(* IEC 61131-3 sources: JingjiangArm/moonboxpro_arm_8.4/Application/Application/任务列表/TensionTask/电机运动/MotionCtl_Trap, 5 files *)

(* ---- StMotorParam_Trap.st ---- *)
(*@CES
Name=StMotorParam_Trap
Type=Gvl
TypeGuid=2db5746d-d284-4425-9f7f-2663a34b0ebc
Guid=895de25e-1961-43a4-b404-7adc5138347b
HasDeclaration=True
HasImplementation=False
*)
{DECLARATION}
TYPE StMotorParam_Trap ://点位轴和龙门轴的参数
STRUCT
	iAxisId: INT;
	iCoreId: INT;
	iStationId: INT;
	iUnitId : INT;
	iMoveStep: INT;
	xMoveRev: BOOL;
	xMoveEn: BOOL;
	uiAxisNum: UINT;(*减速比分子*)
	uiAxisDen: UINT;(*减速比分母*)
	liTargetPos: LINT;(*点位目标位置*)
	udiTargetVel: UDINT;
	rScrewPitch_: REAL;(*螺距*)
END_STRUCT
END_TYPE

{IMPLEMENTATION}

(* ---- KS_FB_AxisPosCtl_Trap.st ---- *)
(*@CES
Name=KS_FB_AxisPosCtl_Trap
Type=FunctionBlock
TypeGuid=6f9dac99-8de1-4efc-8465-68ac443b7d08
Guid=53966cce-5ce5-480b-a4cc-b0ff05bfaf84
HasDeclaration=True
HasImplementation=True
*)
{DECLARATION}
FUNCTION_BLOCK KS_FB_AxisPosCtl_Trap
VAR_INPUT
	i_xEn: BOOL;
	i_iGrpId: INT;
	i_iGrpUnitNum_Pu : INT;
	i_aiGrpUnitList: ARRAY [1..MAX_UNIT_NUM] OF INT;
	i_iGrpTrapMotion_Num: INT;
	i_aiGrpTrapMotion_StdList: ARRAY [1..MAX_STATION_NUM] OF INT;
	i_pstStSysParam: POINTER TO StSysParam;
	i_pastStMotorParam_Trap: POINTER TO ARRAY [1..MAX_STATION_NUM] OF StMotorParam_Trap;

	i_xHorManuCtrl:BOOL;(*界面横向手动修正功能*)

	//2026.01.28.173520 | + | 横向伺服控制
	i_alrTarp_EncPos						: ARRAY [1..MAX_UNIT_NUM] OF LREAL;//横向点位轴的编码器位置
	i_pastStIOMap_AxisBasic					: POINTER TO ARRAY [1..MAX_UNIT_NUM] OF StIOMap_Axis_FE; (*基础io|*)
	i_pastStAxisRapidAdjProf_H				: POINTER TO ARRAY [1..MAX_UNIT_NUM] OF StAxisRapidAdjProf_H;(*纵向快速对版|*)

	i_paxLimit_Left_Wr 						: POINTER TO ARRAY [1..MAX_UNIT_NUM] OF BOOL;
 	i_paxLimit_Right_Wr 					: POINTER TO ARRAY [1..MAX_UNIT_NUM] OF BOOL;
	i_paxLimit_Left_WrClr 					: POINTER TO ARRAY [1..MAX_UNIT_NUM] OF BOOL;
 	i_paxLimit_Right_WrClr 					: POINTER TO ARRAY [1..MAX_UNIT_NUM] OF BOOL;

	//新增拿横向编码器 2026.05.09.104451
	i_pastStGetMotionSts			: POINTER TO ARRAY [1..MAX_STATION_NUM] OF StGetMotionSts;
	i_pstStSysStationInf			:POINTER TO StSysStationInf;
	i_pstStSysGantryAxisInf 		:POINTER TO StSysGantryAxisInf;
	i_pastStAxisIdListInf 			:POINTER TO ARRAY [1..128] OF StAxisIdListInf;
END_VAR
VAR_OUTPUT
END_VAR
VAR
	iN: INT;
	iAxisId: INT;
	iTypeId: INT;
	iUnitId: INT;
	iCoreId: INT;
	pstStGrpParam_Save: POINTER TO StGrpParam_Save;
	pstStGrpParam_UnSave: POINTER TO StGrpParam_UnSave;

	//2026.01.28.173520 | + | 横向伺服控制
	fbKS_FB_HorzCtl_Driver : KS_FB_HorzCtl_Driver;

	alrTotalAdjust_Horz : ARRAY [1..MAX_UNIT_NUM] OF LREAL;
END_VAR

{IMPLEMENTATION}
IF i_xEn THEN
	IF (i_iGrpId=1 OR i_iGrpId=2) AND
		i_iGrpUnitNum_Pu>=1 AND i_iGrpUnitNum_Pu<=MAX_UNIT_NUM AND
		i_iGrpTrapMotion_Num>=1 AND i_iGrpTrapMotion_Num<= MAX_STATION_NUM AND
		i_pstStSysParam<>0 AND
		i_pastStMotorParam_Trap<>0 THEN
		pstStGrpParam_Save:= ADR(i_pstStSysParam^.astStGrpParam_Save[i_iGrpId]);
		pstStGrpParam_UnSave:= ADR(i_pstStSysParam^.astStGrpParam_UnSave[i_iGrpId]);

		//2026.01.28.173520 | + | 横向伺服控制
		fbKS_FB_HorzCtl_Driver(
			i_xEn:= TRUE,//(pstStGrpParam_UnSave^.xFlag_Print OR i_pstStSysParam^.astStGrpParam_Save[i_iGrpId].xEnaTestARC_Ink (*空转测试使能*)) AND g_stStSysParam.stStSysParam_Save.byHorzCtlMode=3,
			i_iGrpId:= i_iGrpId,
			i_iGrpAxisNum_Pu:= i_iGrpUnitNum_Pu,
			i_pstStSysParam:= i_pstStSysParam,
			i_pastStIOMap_AxisBasic:= i_pastStIOMap_AxisBasic,
			i_lrVel_HorzAdjust:= REAL_TO_LREAL(i_pstStSysParam^.astStGrpParam_Save[i_iGrpId].rVel_HorzdAdj),
			i_lrVel_HorzPreRegister:=  REAL_TO_LREAL(i_pstStSysParam^.astStGrpParam_Save[i_iGrpId].rVel_HorzPreRegister),
			i_xFlag_Estop:= pstStGrpParam_UnSave^.xFlag_EStop,
			i_xFlag_Stop:= pstStGrpParam_UnSave^.xFlag_Stop,
			i_iCycleTime_Plc:= gc_TENSION_TSK_CYCLE_TIME,
			i_pastStAxisRapidAdjProf_H:= i_pastStAxisRapidAdjProf_H,
			i_alrTarp_EncPos:= i_alrTarp_EncPos,
			i_paxLimit_Left_Wr:= i_paxLimit_Left_Wr,
			i_paxLimit_Right_Wr:= i_paxLimit_Right_Wr,
			i_paxLimit_Left_WrClr:= i_paxLimit_Left_WrClr,
			i_paxLimit_Right_WrClr:= i_paxLimit_Right_WrClr,
			i_xHorManuCtrl:= i_xHorManuCtrl,
			i_aiGrpTrapMotion_StdList:=i_aiGrpTrapMotion_StdList,
			i_pastStGetMotionSts:=i_pastStGetMotionSts,
			i_pstStSysStationInf:=i_pstStSysStationInf,
			i_pstStSysGantryAxisInf :=i_pstStSysGantryAxisInf,
			i_pastStAxisIdListInf :=i_pastStAxisIdListInf,
			o_xEno=> ,
			o_iErNo=> ,
			o_alrTotalAdjust_Horz=> alrTotalAdjust_Horz);

		FOR iN:=1 TO i_iGrpTrapMotion_Num BY 1 DO
			i_pastStMotorParam_Trap^[iN].liTargetPos := LREAL_TO_LINT(alrTotalAdjust_Horz[iN]*
						i_pstStSysParam^.astStUnitParam_Save[iN].uiNum_Horz*
						GC_LRMOTORPPR_TRAP/
						i_pstStSysParam^.astStUnitParam_Save[iN].rScrewPitch_Horz/
						i_pstStSysParam^.astStUnitParam_Save[iN].uiDen_Horz/1000.0);
			i_pastStMotorParam_Trap^[iN].udiTargetVel := LREAL_TO_UDINT(i_pstStSysParam^.astStGrpParam_Save[i_iGrpId].rVel_HorzdAdj*
						i_pstStSysParam^.astStUnitParam_Save[iN].uiNum_Horz*
						GC_LRMOTORPPR_TRAP/
						i_pstStSysParam^.astStUnitParam_Save[iN].rScrewPitch_Horz/
						i_pstStSysParam^.astStUnitParam_Save[iN].uiDen_Horz/1000.0);
		END_FOR
	END_IF
ELSE
	;
END_IF

(* ---- KS_FB_HorzCtl_Driver.st ---- *)
(*@CES
Name=KS_FB_HorzCtl_Driver
Type=FunctionBlock
TypeGuid=6f9dac99-8de1-4efc-8465-68ac443b7d08
Guid=da6152f2-d53e-407a-9477-cd718a7d485f
HasDeclaration=True
HasImplementation=True
*)
{DECLARATION}
FUNCTION_BLOCK KS_FB_HorzCtl_Driver
VAR_INPUT
	i_xEn: BOOL;(*使能*)
	i_iGrpId: INT;
	i_iGrpAxisNum_Pu: INT; (*色组轴数*)
	i_pstStSysParam:POINTER TO StSysParam;(*系参数*)
	i_pastStIOMap_AxisBasic					: POINTER TO ARRAY [1..MAX_UNIT_NUM] OF StIOMap_Axis_FE; (*基础io|*)
	i_lrVel_HorzAdjust		: LREAL;(*mm/s; um/ms; 横向调整速度|*)
	i_lrVel_HorzPreRegister		: LREAL;(*mm/s;横向预套准速度|*)
	(*2023.3.8.114628*)
	i_xFlag_Estop							: BOOL;(*急停标志*)
	i_xFlag_Stop							: BOOL;(*停机标志*)
	i_iCycleTime_Plc						: INT;
	i_pastStAxisRapidAdjProf_H				: POINTER TO ARRAY [1..MAX_UNIT_NUM] OF StAxisRapidAdjProf_H;(*纵向快速对版|*)
	i_alrTarp_EncPos						: ARRAY [1..MAX_UNIT_NUM] OF LREAL;//横向点位轴的编码器位置
	i_paxLimit_Left_Wr 						: POINTER TO ARRAY [1..MAX_UNIT_NUM] OF BOOL;
 	i_paxLimit_Right_Wr 					: POINTER TO ARRAY [1..MAX_UNIT_NUM] OF BOOL;
	i_paxLimit_Left_WrClr 						: POINTER TO ARRAY [1..MAX_UNIT_NUM] OF BOOL;
 	i_paxLimit_Right_WrClr 					: POINTER TO ARRAY [1..MAX_UNIT_NUM] OF BOOL;
	i_xHorManuCtrl:BOOL;(*界面横向手动修正功能*)
//	i_arStep_Horz			:POINTER TO ARRAY [1..MAX_UNIT_NUM] OF REAL;
//2026.05.09.100428 新增横向标定功能
	i_aiGrpTrapMotion_StdList: ARRAY [1..MAX_STATION_NUM] OF INT;
	i_pastStGetMotionSts: POINTER TO ARRAY [1..MAX_STATION_NUM] OF StGetMotionSts;
	i_pstStSysStationInf			:POINTER TO StSysStationInf;
	i_pstStSysGantryAxisInf 		:POINTER TO StSysGantryAxisInf;
	i_pastStAxisIdListInf :POINTER TO ARRAY [1..128] OF StAxisIdListInf;
END_VAR
VAR_OUTPUT
	o_xEno: BOOL;
	o_iErNo: INT;(*0成功\-1参数失败|*)
	o_alrTotalAdjust_Horz: ARRAY [1..MAX_UNIT_NUM] OF LREAL;(*横向调整量*)

END_VAR
VAR
	iN: INT;
	xInit: BOOL;
	iAxisId: INT;
	pstStGrpParam_Save: POINTER TO StGrpParam_Save;
	pstStGrpParam_UnSave: POINTER TO StGrpParam_UnSave;

	pstStUnitParam_Save: POINTER TO StUnitParam_Save;
	pstStUnitParam_UnSave: POINTER TO StUnitParam_UnSave;
	pstStRSV_UnitParam_Save: POINTER TO StRSV_UnitParam_Save;
	pstStRSV_UnitParam_UnSave: POINTER TO StRSV_UnitParam_UnSave;
	(*横向运动相关变量都使用操作侧和传动侧变量重新赋值@2023.3.8.104853*)
	axHorMovingBtn_M: ARRAY [1..MAX_UNIT_NUM] OF BOOL;(*横向操作侧运动按钮*)
	axHorMovingBtn_G: ARRAY [1..MAX_UNIT_NUM] OF BOOL;(*横向传动侧运动按钮*)
	axHorMovingLimit_M: ARRAY [1..MAX_UNIT_NUM] OF BOOL;(*横向操作侧运动限位*)
	axHorMovingLimit_G: ARRAY [1..MAX_UNIT_NUM] OF BOOL;(*横向传动侧运动限位*)
	axHorMoving_M: ARRAY [1..MAX_UNIT_NUM] OF BOOL;(*横向操作侧运动*)
	axHorMoving_G: ARRAY [1..MAX_UNIT_NUM] OF BOOL;(*横向传动侧运动*)

	lrAdjustVel_:LREAL;(*每个周期调整的量|这里还是mm/s，需要转化为*)
	alrTotalAdjust_Horz: ARRAY [1..MAX_UNIT_NUM] OF LREAL;(*横向调整量*)
	adwTotalTimes_CW_AxisHorzManu: ARRAY [1..MAX_UNIT_NUM] OF DWORD := [MAX_UNIT_NUM(0)];
	adwTotalTimes_CCW_AxisHorzManu: ARRAY [1..MAX_UNIT_NUM] OF DWORD := [MAX_UNIT_NUM(0)];

	wHorzMotorDir: WORD;(*.0 |正转方向
					.1|反转方向*)
	awPreHorzMotorDir: ARRAY [1..MAX_UNIT_NUM] OF WORD;
	axHorzMotorStart_Delay: ARRAY [1..MAX_UNIT_NUM] OF BOOL;(*横向启动延时标志*)
	axHorzMotorStart_DelayDne: ARRAY [1..MAX_UNIT_NUM] OF BOOL;(*横向启动延时完成*)
	auiHorzMotorStart_Count: ARRAY [1..MAX_UNIT_NUM] OF UINT;(*启动延时计时变量*)
	iHorzMotorStart_DelayTime_MS: INT:=0;(*启动的延时时间ms*)

	axStopManuMove_Horz: ARRAY  [1..MAX_UNIT_NUM] OF BOOL;
	lrLimit_Left:LREAL;
	lrLimit_Right:LREAL;
	xLimit_LeftTemp:BOOL;
	xLimit_RightTemp:BOOL;
	xLimit_Left:BOOL;
	xLimit_Right:BOOL;
	lrAbsPosHorz:LREAL;
	iRtn:INT;
	xAxisRev:BOOL;

	//2026.05.09.170157 | + | 增加正反流向
	xMachineIsRev : BOOL;
END_VAR

{IMPLEMENTATION}
o_xEno:= i_xEn;
o_iErNo:= 0;
IF i_xEn THEN
	IF (i_iGrpAxisNum_Pu>=1 AND i_iGrpAxisNum_Pu<=MAX_UNIT_NUM) AND(*系的色组数量有效|*)
		i_pstStSysParam<>0 AND(*参数有效|*)
		i_pastStIOMap_AxisBasic<>0 AND
		i_paxLimit_Left_Wr<>0 AND
		i_paxLimit_Right_Wr<>0 THEN

		pstStGrpParam_Save :=  ADR(i_pstStSysParam^.astStGrpParam_Save[i_iGrpId]);
		pstStGrpParam_UnSave :=  ADR(i_pstStSysParam^.astStGrpParam_UnSave[i_iGrpId]);
		//初始化输出调整量为当前规划位置
// 		IF NOT xInit THEN
// 			xInit:= TRUE;
// 			FOR iN:=1 TO i_iGrpAxisNum_Pu BY 1 DO
// 				alrTotalAdjust_Horz[iN]:= i_alrTarp_PrfPos[iN];
// 			END_FOR
// 		END_IF

		//2026.05.09.170157 | + | 增加正反流向
		xMachineIsRev := TRUE;

		IF NOT xInit THEN
			xInit:= TRUE;
			FOR iN:=1 TO i_iGrpAxisNum_Pu BY 1 DO
				alrTotalAdjust_Horz[iN]:= 0;
			END_FOR
		END_IF
		(*2023.3.8.114227 将函数KS_FB_AxisHorAdj中的代码移植到此处*)
		FOR iN:= 1 TO i_iGrpAxisNum_Pu BY 1 DO
			iAxisId:= iN;
			pstStUnitParam_Save:= ADR(i_pstStSysParam^.astStUnitParam_Save[iAxisId]);
			pstStUnitParam_UnSave:= ADR(i_pstStSysParam^.astStUnitParam_UnSave[iAxisId]);

			pstStRSV_UnitParam_Save := ADR(i_pstStSysParam^.astStRSV_UnitParam_Save[iAxisId]);
			pstStRSV_UnitParam_UnSave := ADR(i_pstStSysParam^.astStRSV_UnitParam_UnSave[iAxisId]);

			(*处理一下限位*)
			(*限位赋值*)
			IF pstStGrpParam_UnSave^.xIsDebugMode_Machine AND pstStGrpParam_UnSave^.xFlag_Stop THEN//调试模式
				//记录一下横向限位
				IF i_paxLimit_Left_Wr^[iAxisId] THEN
					i_paxLimit_Left_Wr^[iAxisId]:= FALSE;
					//2026.05.09.100428 新增横向标定功能 Hou.N
					iRtn := GTN_RN_ReadAbsEncPos(cardIndex:= 1, stationPhyId:=i_aiGrpTrapMotion_StdList[iAxisId], encoder:= 1, pPos:= ADR(lrAbsPosHorz));
					g_liAbsPosTrap := LREAL_TO_LINT(lrAbsPosHorz);
					xAxisRev := pstStUnitParam_UnSave^.xMotRev_Horiz_;
					iRtn := KS_SetTrapCoordinate(
							i_xEn:= TRUE,
							i_iTarget_Num:= 1,
							i_paiTargetStationList:= ADR(i_aiGrpTrapMotion_StdList[iAxisId]),
							i_paliABSEncPos:= ADR(g_liAbsPosTrap),
							i_paxAxisRev:= ADR(xAxisRev),
							i_pastStAxisIdListInf:= i_pastStAxisIdListInf,
							i_pastStGetMotionSts:= i_pastStGetMotionSts,
							i_pstStSysStationInf := i_pstStSysStationInf,
							i_pstStSysGantryAxisInf := i_pstStSysGantryAxisInf,
							ADR(g_alrCurrentAbsPos_Trap));
					i_pstStSysParam^.astStRSV_UnitParam_Save[iAxisId].liABSPos_Trap:= g_liAbsPosTrap;
					pstStRSV_UnitParam_Save^.lrLimit_Left:= 1;
				END_IF

				IF i_paxLimit_Right_Wr^[iAxisId] THEN
					i_paxLimit_Right_Wr^[iAxisId]:= FALSE;
					pstStRSV_UnitParam_Save^.lrLimit_Right:= i_alrTarp_EncPos[iAxisId];
				END_IF
				IF 	i_paxLimit_Left_WrClr^[iAxisId] THEN
					i_paxLimit_Left_WrClr^[iAxisId] := FALSE;
					pstStRSV_UnitParam_Save^.lrLimit_Left := 0;
					i_pstStSysParam^.astStRSV_UnitParam_Save[iAxisId].liABSPos_Trap:=0;
				END_IF
				IF 	i_paxLimit_Right_WrClr^[iAxisId] THEN
					i_paxLimit_Right_WrClr^[iAxisId] := FALSE;
					pstStRSV_UnitParam_Save^.lrLimit_Right := 0;
				END_IF
			ELSE
				i_paxLimit_Left_Wr^[iAxisId]:= FALSE;
				i_paxLimit_Right_Wr^[iAxisId]:= FALSE;
				i_paxLimit_Left_WrClr^[iAxisId]:= FALSE;
				i_paxLimit_Right_WrClr^[iAxisId]:= FALSE;
			END_IF
			lrLimit_Left:= pstStRSV_UnitParam_Save^.lrLimit_Left;
			lrLimit_Right:= pstStRSV_UnitParam_Save^.lrLimit_Right;
			xLimit_LeftTemp:=i_pastStIOMap_AxisBasic^[iAxisId].i_xPosLimit_Left;
			xLimit_RightTemp:=i_pastStIOMap_AxisBasic^[iAxisId].i_xPosLimit_Right;

			IF lrLimit_Left=0 THEN(*未有软限位|按照最远距离*);

			ELSE(*存在软限位|限位标志取接近开关和位置值的or*)
				IF pstStUnitParam_UnSave^.xMotRev_Horiz_ THEN
					xLimit_LeftTemp:=xLimit_LeftTemp OR
									(lrLimit_Left<i_alrTarp_EncPos[iAxisId]);
				ELSE
					xLimit_LeftTemp:=xLimit_LeftTemp OR
									(lrLimit_Left<i_alrTarp_EncPos[iAxisId]);
				END_IF
			END_IF
			IF lrLimit_Right=0 THEN(*未有软限位|按照最远距离*);
			ELSE(*存在软限位|限位标志取接近开关和位置值的or*)
				IF pstStUnitParam_UnSave^.xMotRev_Horiz_ THEN
					xLimit_RightTemp:=xLimit_RightTemp OR
								(lrLimit_Right>i_alrTarp_EncPos[iAxisId]);
				ELSE
					xLimit_RightTemp:=xLimit_RightTemp OR
								(lrLimit_Right>i_alrTarp_EncPos[iAxisId]);

				END_IF
			END_IF

			(*手动左右取反*)(*bai.zy|2023.12.18.161830|feida取反*)
			xLimit_Left:=xLimit_RightTemp;
			xLimit_Right:=xLimit_LeftTemp;
			(*
			IF xMachineIsRev THEN
				xLimit_Left:=xLimit_RightTemp;
				xLimit_Right:=xLimit_LeftTemp;
				IF pstStUnitParam_UnSave^.xMotRev_Horiz_ THEN
					xLimit_Left:=xLimit_LeftTemp;
					xLimit_Right:=xLimit_RightTemp;
				END_IF
			ELSE
				xLimit_Left:=xLimit_LeftTemp;
				xLimit_Right:=xLimit_RightTemp;
				IF pstStUnitParam_UnSave^.xMotRev_Horiz_ THEN
					xLimit_Left:=xLimit_LeftTemp;
					xLimit_Right:=xLimit_RightTemp;
				END_IF
			END_IF
			*)
//2026.01.28.152311 | + | 界面上的限位提示，先不要了
// 			g_axLimit_Left_Wr_HMI[iN]:= xLimit_Left;
// 			g_axLimit_Right_Wr_HMI[iN]:= xLimit_Right;
			(*处理横向开关相关@2023.3.8.104924*)
			(*和运动方向关联@伺服正转(正手机)-左对应操作侧#先不关心反印时候的方向变化问题
						    @伺服反转(反手机)-左对应传动侧#先不关心反印时候的方向变化问题*)

//			IF pstStUnitParam^.xMotRev_PrnRoller THEN(*正转*)
				axHorMovingBtn_M[iAxisId]:=i_pastStIOMap_AxisBasic^[iAxisId].i_xMove_Left;
				axHorMovingBtn_G[iAxisId]:=i_pastStIOMap_AxisBasic^[iAxisId].i_xMove_Right;

				axHorMovingLimit_M[iAxisId]:=xLimit_Left;
				axHorMovingLimit_G[iAxisId]:=xLimit_Right;
(*			ELSE(*反转*)
				axHorMovingBtn_M[iAxisId]:=pstStIOMap_Axis_FLEXO^.i_xMove_Right;
				axHorMovingBtn_G[iAxisId]:=pstStIOMap_Axis_FLEXO^.i_xMove_Left;

				IF i_pstStSysParam^.dwControlComplexBits.17 THEN
					(*使用左右限位*)
					axHorMovingLimit_M[iAxisId]:=xLimit_Right;
					axHorMovingLimit_G[iAxisId]:=xLimit_Left;
				ELSE
					(*使用正转(操作侧)反转(传动侧)限位*)
					axHorMovingLimit_M[iAxisId]:=xLimit_Left;
					axHorMovingLimit_G[iAxisId]:=xLimit_Right;
				END_IF
			END_IF
*)

			IF i_pastStIOMap_AxisBasic^[iAxisId].o_xRel_Press OR (NOT i_pastStIOMap_AxisBasic^[iAxisId].i_xHorzMotor_FastSpd) THEN
			(*快调/慢调处理*)
				lrAdjustVel_:= i_lrVel_HorzAdjust;
			ELSE
				lrAdjustVel_:= i_lrVel_HorzPreRegister;
			END_IF

			(*2019.5.15.170941|niu.j|急停清零横向调整量*)
			IF pstStGrpParam_UnSave^.xFlag_EStoping OR pstStGrpParam_UnSave^.xFlag_Estop THEN
				pstStUnitParam_UnSave^.alrTotalAdjustVal_Auto_vh[2]:= 0;
				pstStUnitParam_UnSave^.alrTotalAdjustVal_ManuFine_vh[2]:= 0;
				pstStUnitParam_UnSave^.alrTotalAdjustVal_Rapid_vh[2]:= 0;
			END_IF

			IF (pstStUnitParam_Save^.dwFlag_Ctl.0 AND pstStUnitParam_Save^.dwFlag_Sts.1) THEN
				IF ABS(pstStUnitParam_UnSave^.alrTotalAdjustVal_Auto_vh[2])>0 THEN
					IF pstStUnitParam_UnSave^.alrTotalAdjustVal_Auto_vh[2]>0 THEN
						(*正向*)
						alrTotalAdjust_Horz[iAxisId]:= alrTotalAdjust_Horz[iAxisId]+pstStUnitParam_UnSave^.alrTotalAdjustVal_Auto_vh[2];
						pstStUnitParam_UnSave^.alrTotalAdjustVal_Auto_vh[2]:= 0;
						pstStUnitParam_UnSave^.axCurCycleAdjustVal_Auto_done_vh[2]:= FALSE;
						axHorMoving_M[iAxisId]:= TRUE;(*操作侧*)
						axHorMoving_G[iAxisId]:= FALSE;(*传动侧*)
					ELSE
						(*反向*)
						alrTotalAdjust_Horz[iAxisId]:= alrTotalAdjust_Horz[iAxisId]+pstStUnitParam_UnSave^.alrTotalAdjustVal_Auto_vh[2];
						pstStUnitParam_UnSave^.alrTotalAdjustVal_Auto_vh[2]:= 0;
						pstStUnitParam_UnSave^.axCurCycleAdjustVal_Auto_done_vh[2]:= FALSE;
						axHorMoving_G[iAxisId]:= TRUE;(*传动侧*)
						axHorMoving_M[iAxisId]:= FALSE;(*操作侧*)
					END_IF
				ELSE
					IF pstStUnitParam_UnSave^.xFlag_HorzPreRegister_ing THEN
						pstStUnitParam_UnSave^.alrTotalAdjustVal_Auto_vh[2]:= 0;
					END_IF
					axHorMoving_M[iAxisId]:= FALSE;
					axHorMoving_G[iAxisId]:= FALSE;
				END_IF
			ELSIF i_xHorManuCtrl THEN//i_pstStSysParam^.dwControlComplexBits.7 THEN(*界面上有横向手动修正功能|*)
				(*消耗手动细调量累计|*)
				IF ABS(pstStUnitParam_UnSave^.alrTotalAdjustVal_ManuFine_vh[2])>0 THEN
(*					IF axHorzMotorStart_DelayDne[iAxisId] THEN(*延时启动完成了*)
*)						IF pstStUnitParam_UnSave^.alrTotalAdjustVal_ManuFine_vh[2]>0 THEN
							(*正向*)
							alrTotalAdjust_Horz[iAxisId]:= alrTotalAdjust_Horz[iAxisId]+pstStUnitParam_UnSave^.alrTotalAdjustVal_ManuFine_vh[2];
							pstStUnitParam_UnSave^.alrTotalAdjustVal_ManuFine_vh[2]:= 0;
							pstStUnitParam_UnSave^.axCurCycleAdjustVal_ManuFine_done_vh[2]:= FALSE;
							axHorMoving_M[iAxisId]:= TRUE;(*操作侧*)
							axHorMoving_G[iAxisId]:= FALSE;(*传动侧*)

						ELSE
							(*反向*)
							alrTotalAdjust_Horz[iAxisId]:= alrTotalAdjust_Horz[iAxisId]+pstStUnitParam_UnSave^.alrTotalAdjustVal_ManuFine_vh[2];
							pstStUnitParam_UnSave^.alrTotalAdjustVal_ManuFine_vh[2]:= 0;
							pstStUnitParam_UnSave^.axCurCycleAdjustVal_ManuFine_done_vh[2]:= FALSE;
							axHorMoving_G[iAxisId]:= TRUE;(*传动侧*)
							axHorMoving_M[iAxisId]:= FALSE;(*操作侧*)

						END_IF

					(*monitoring...\2018.10.7.104410|*)
					IF axHorMoving_M[iAxisId] THEN
						adwTotalTimes_CW_AxisHorzManu[iAxisId]:= adwTotalTimes_CW_AxisHorzManu[iAxisId]+1;
					END_IF
					IF axHorMoving_G[iAxisId] THEN
						adwTotalTimes_CCW_AxisHorzManu[iAxisId]:= adwTotalTimes_CCW_AxisHorzManu[iAxisId]+1;
					END_IF

				ELSE
					axHorMoving_M[iAxisId]:= FALSE;
					axHorMoving_G[iAxisId]:= FALSE;
				END_IF
			ELSE
				(*没开横向或者横向在手动状态*)
				pstStUnitParam_UnSave^.axCurCycleAdjustVal_Auto_done_vh[2]:= FALSE;
				pstStUnitParam_UnSave^.axCurCycleAdjustVal_Rapid_done_vh[2]:= FALSE;
				pstStUnitParam_UnSave^.axCurCycleAdjustVal_ManuCoarse_done_vh[2]:= FALSE;
				pstStUnitParam_UnSave^.axCurCycleAdjustVal_ManuFine_done_vh[2]:= FALSE;
				pstStUnitParam_UnSave^.axCurCycleAdjustVal_Coupling_done_vh[2]:= FALSE;
//				pstStUnitParam^.axCurCycleAdjustVal_Compensate_done_vh[2]:= FALSE;

				pstStUnitParam_UnSave^.alrCurCycleAdjustVal_Auto_vh[2]:= 0;
				pstStUnitParam_UnSave^.alrCurCycleAdjustVal_Rapid_vh[2]:= 0;
				pstStUnitParam_UnSave^.alrCurCycleAdjustVal_ManuCoarse_vh[2]:= 0;
				pstStUnitParam_UnSave^.alrCurCycleAdjustVal_ManuFine_vh[2]:= 0;
				pstStUnitParam_UnSave^.alrCurCycleAdjustVal_Coupling_vh[2]:= 0;
//				pstStUnitParam^.alrCurCycleAdjustVal_Compensate_vh[2]:= 0;

				pstStUnitParam_UnSave^.alrTotalAdjustVal_Auto_vh[2]:= 0;
				pstStUnitParam_UnSave^.alrTotalAdjustVal_Rapid_vh[2]:= 0;
(*				pstStUnitParam^.alrTotalAdjustVal_ManuCoarse_vh[2]:= 0;*)
				pstStUnitParam_UnSave^.alrTotalAdjustVal_ManuFine_vh[2]:= 0;
				pstStUnitParam_UnSave^.alrTotalAdjustVal_Coupling_vh[2]:= 0;
//				pstStUnitParam^.alrTotalAdjustVal_Compensate_vh[2]:= 0;

				axHorMoving_M[iAxisId]:= FALSE;
				axHorMoving_G[iAxisId]:= FALSE;
			END_IF

			(*增加了正反转信号启动延时2018.10.7.085705 by liu.yt*)
			wHorzMotorDir:=BOOL_TO_WORD(axHorMoving_M[iAxisId])+SHL(BOOL_TO_WORD(axHorMoving_G[iAxisId]),1);
			IF wHorzMotorDir<>awPreHorzMotorDir[iAxisId] THEN(*方向发生了变化*)
				IF wHorzMotorDir<>0THEN(*说明有正反转信号了*)
					axHorzMotorStart_Delay[iAxisId]:=TRUE;
				ELSE
					axHorzMotorStart_Delay[iAxisId]:=FALSE;
				END_IF
				axHorzMotorStart_DelayDne[iAxisId]:=FALSE;
				auiHorzMotorStart_Count[iAxisId]:=0;
				awPreHorzMotorDir[iAxisId]:=wHorzMotorDir;
			END_IF

			IF axHorzMotorStart_Delay[iAxisId] THEN(*启动延时*)
				IF auiHorzMotorStart_Count[iAxisId]>=iHorzMotorStart_DelayTime_MS/i_iCycleTime_Plc THEN
					auiHorzMotorStart_Count[iAxisId]:=0;
					axHorzMotorStart_Delay[iAxisId]:=FALSE;
					axHorzMotorStart_DelayDne[iAxisId]:=TRUE;
				ELSE
					auiHorzMotorStart_Count[iAxisId]:=auiHorzMotorStart_Count[iAxisId]+1;
				END_IF
			END_IF

			IF i_pstStSysParam^.astStRSV_UnitParam_UnSave[iAxisId].xBtn_FromHMI_HorMove_M THEN
				i_pstStSysParam^.astStRSV_UnitParam_UnSave[iAxisId].xBtn_FromHMI_HorMove_G:= FALSE;
				i_pstStSysParam^.astStRSV_UnitParam_UnSave[iAxisId].xBtn_FromHMI_HorMove_M:= FALSE;
				IF NOT xLimit_Left THEN
					alrTotalAdjust_Horz[iAxisId]:= alrTotalAdjust_Horz[iAxisId]-
						REAL_TO_LREAL(i_pstStSysParam^.astStRSV_UnitParam_UnSave[iAxisId].rStep_Horz*1000.0);
				END_IF
			ELSIF i_pstStSysParam^.astStRSV_UnitParam_UnSave[iAxisId].xBtn_FromHMI_HorMove_G THEN
				i_pstStSysParam^.astStRSV_UnitParam_UnSave[iAxisId].xBtn_FromHMI_HorMove_M:= FALSE;
				i_pstStSysParam^.astStRSV_UnitParam_UnSave[iAxisId].xBtn_FromHMI_HorMove_G:= FALSE;
				IF NOT xLimit_Right THEN
					alrTotalAdjust_Horz[iAxisId]:= alrTotalAdjust_Horz[iAxisId]+
						REAL_TO_LREAL(i_pstStSysParam^.astStRSV_UnitParam_UnSave[iAxisId].rStep_Horz*1000.0);
				END_IF
			END_IF
// 			(*2026.2.10.095914 增加从站横向步进量调整*)
// 			IF pstStRSV_UnitParam_UnSave^.xHorMoving_M AND (NOT pstStRSV_UnitParam_UnSave^.xHorMoving_G) AND (NOT xLimit_Left) THEN
// 				(*左*)
// 				alrTotalAdjust_Horz[iAxisId]:= alrTotalAdjust_Horz[iAxisId]-REAL_TO_LREAL(pstStRSV_UnitParam_UnSave^.rStep_Horz)
// 				;
// 				axHorMoving_G[iAxisId]:= FALSE;
// 				axHorMoving_M[iAxisId]:= TRUE;
//
// 			ELSIF pstStRSV_UnitParam_UnSave^.xHorMoving_G AND (NOT pstStRSV_UnitParam_UnSave^.xHorMoving_M) AND (NOT xLimit_Right) THEN
// 				(*右*)
// 				alrTotalAdjust_Horz[iAxisId]:= alrTotalAdjust_Horz[iAxisId]+REAL_TO_LREAL(pstStRSV_UnitParam_UnSave^.rStep_Horz)
// 				;
// 				axHorMoving_M[iAxisId]:= FALSE;
// 				axHorMoving_G[iAxisId]:= TRUE;
// 			ELSE
// 				axHorMoving_M[iAxisId]:= FALSE;
// 				axHorMoving_G[iAxisId]:= FALSE;
// 			END_IF
//

			(*---------------------------2017-08-14 15:21:18
			/.手动调整
			.----------------------------------------------*)
			IF axHorMovingBtn_M[iAxisId]  AND (NOT axHorMovingBtn_G[iAxisId]) AND (NOT xLimit_Left) (*AND
			(NOT pstStRSV_UnitParam_UnSave^.xHorMoving_G)	AND
			(NOT pstStRSV_UnitParam_UnSave^.xHorMoving_M)*) THEN
				(*左*)
				alrTotalAdjust_Horz[iAxisId]:= alrTotalAdjust_Horz[iAxisId]-
				i_lrVel_HorzAdjust*	i_iCycleTime_Plc*1;

				axHorMoving_G[iAxisId]:= FALSE;
				axHorMoving_M[iAxisId]:= TRUE;
			ELSIF axHorMovingBtn_G[iAxisId]  AND (NOT axHorMovingBtn_M[iAxisId]) AND (NOT xLimit_Right)(* AND
			(NOT pstStRSV_UnitParam_UnSave^.xHorMoving_G)	AND
			(NOT pstStRSV_UnitParam_UnSave^.xHorMoving_M) *) THEN
				(*右*)
				alrTotalAdjust_Horz[iAxisId]:= alrTotalAdjust_Horz[iAxisId]+
				i_lrVel_HorzAdjust*	i_iCycleTime_Plc*1;

				axHorMoving_M[iAxisId]:= FALSE;
				axHorMoving_G[iAxisId]:= TRUE;
			ELSE

				axHorMoving_M[iAxisId]:= FALSE;
				axHorMoving_G[iAxisId]:= FALSE;

// 			ELSIF (NOT  axHorMovingBtn_G[iAxisId])  AND
// 				(NOT axHorMovingBtn_M[iAxisId]) AND
// 				(NOT axStopManuMove_Horz[iAxisId]) THEN
// 				axStopManuMove_Horz[iAxisId]:= TRUE;
// 				axHorMoving_M[iAxisId]:= FALSE;
// 				axHorMoving_G[iAxisId]:= FALSE;
// 				alrTotalAdjust_Horz[iAxisId]:= i_alrTarp_PrfPos[iAxisId]*
// 						pstStUnitParam^.uiDen_Horz*1000.0*pstStUnitParam^.rScrewPitch_Horz/
// 						GC_LRMOTORPPR_TRAP/UINT_TO_LREAL(pstStUnitParam^.uiNum_Horz);
// 				IF pstStUnitParam^.xMotRev_Horiz_ THEN
// 					alrTotalAdjust_Horz[iAxisId]:= -alrTotalAdjust_Horz[iAxisId];
// 				END_IF
			END_IF

			(*---------------------------2017-08-14 15:21:18
			/.横向限位处理
			.----------------------------------------------*)
			IF axHorMovingLimit_M[iAxisId] THEN(*操作侧*)
				axHorMoving_M[iAxisId]:= FALSE;
			END_IF

			IF axHorMovingLimit_G[iAxisId] THEN(*传动侧*)
				axHorMoving_G[iAxisId]:= FALSE;
			END_IF

			(*急停停止横向输出|2022.5.11.171513*)
			IF pstStGrpParam_UnSave^.xFlag_EStoping OR pstStGrpParam_UnSave^.xFlag_Estop THEN
				axHorMoving_M[iAxisId]:= FALSE;
				axHorMoving_G[iAxisId]:= FALSE;
			END_IF

			(*将操作侧和传动侧信号输出*)
			(*电机输出是按照正转和反转@一般情况正反手机电机的旋转方向是一致的即,都是向操作侧或者都是向传动侧
			我们定义正传是向操作侧@反转是向传动侧*)
//2026.5.12.143337点位控制横向不需要再输出到IO了
// 			i_pastStIOMap_AxisBasic^[iAxisId].o_xHorzMotor_CW:=axHorMoving_M[iAxisId];
// 			i_pastStIOMap_AxisBasic^[iAxisId].o_xHorzMotor_CCW:=axHorMoving_G[iAxisId];
			//2023.9.25.174830确定输出方向
			o_alrTotalAdjust_Horz[iAxisId]:= alrTotalAdjust_Horz[iAxisId];
			IF pstStUnitParam_UnSave^.xMotRev_Horiz_ THEN
				o_alrTotalAdjust_Horz[iAxisId]:= -o_alrTotalAdjust_Horz[iAxisId];
			END_IF
		END_FOR
	END_IF
END_IF

(* ---- KS_FB_MotionCtl_Trap.st ---- *)
(*@CES
Name=KS_FB_MotionCtl_Trap
Type=FunctionBlock
TypeGuid=6f9dac99-8de1-4efc-8465-68ac443b7d08
Guid=91bb1670-7a0e-427e-a57a-b27b647b87fa
HasDeclaration=True
HasImplementation=True
*)
{DECLARATION}
FUNCTION_BLOCK KS_FB_MotionCtl_Trap
VAR_INPUT
	i_xEn: BOOL;
	i_iGrpId: INT;
	i_iGrpUnitNum_Pu : INT;
	i_aiGrpUnitList: ARRAY [1..MAX_UNIT_NUM] OF INT;
	i_iGrpTrapMotion_Num: INT;
	i_aiGrpTrapMotion_StdList: ARRAY [1..MAX_STATION_NUM] OF INT;

	i_pstStSysParam: POINTER TO StSysParam;
	i_pastStSetPrm					:POINTER TO ARRAY [1..MAX_STATION_NUM] OF TSetMultiMcFunctionPrm;
	i_pastStGetMotionSts: POINTER TO ARRAY [1..MAX_STATION_NUM] OF StGetMotionSts;
	i_pastStMotorParam_Trap: POINTER TO ARRAY [1..MAX_STATION_NUM] OF StMotorParam_Trap;
	i_pstStHYLogFifo			: POINTER TO StHYLogFifo;(* 2025.8.23.170701/han.dp/增加的日志队列 *)
	i_pastStIOMap_Main_FE						: POINTER TO ARRAY [1..4] OF StIOMap_Main_FE;(*轴io数据区域|AB系*)
	i_pastStIOMap_Axis_FE					: POINTER TO ARRAY [1..MAX_UNIT_NUM] OF StIOMap_Axis_FE;(*轴io数据区域|*)
	i_pstStSysStationInf			:POINTER TO StSysStationInf;
	i_pstStSysGantryAxisInf : POINTER TO StSysGantryAxisInf;

	i_xHorManuCtrl:BOOL;(*界面横向手动修正功能*)
	i_pastStAxisRapidAdjProf_H				: POINTER TO ARRAY [1..MAX_UNIT_NUM] OF StAxisRapidAdjProf_H;(*纵向快速对版|*)

	i_paxLimit_Left_Wr 						: POINTER TO ARRAY [1..MAX_UNIT_NUM] OF BOOL;
 	i_paxLimit_Right_Wr 					: POINTER TO ARRAY [1..MAX_UNIT_NUM] OF BOOL;
	i_paxLimit_Left_WrClr 					: POINTER TO ARRAY [1..MAX_UNIT_NUM] OF BOOL;
 	i_paxLimit_Right_WrClr 					: POINTER TO ARRAY [1..MAX_UNIT_NUM] OF BOOL;
	i_pastStAxisIdListInf 			:POINTER TO ARRAY [1..128] OF StAxisIdListInf;
END_VAR
VAR_OUTPUT
END_VAR
VAR_IN_OUT
END_VAR
VAR
	pstStGrpParam_Save : POINTER TO StGrpParam_Save;
	pstStGrpParam_UnSave : POINTER TO StGrpParam_UnSave;

	dwRtn : DWORD;
	iRtn : INT;
	astStSetPrm_Pre				: ARRAY [1..MAX_STATION_NUM] OF TSetMultiMcFunctionPrm;
	stStGetPrm				: TMultiMcFunctionReadPrm;
	iMaxRetryTimes: INT := 3;
	aiRetryCount: ARRAY [1..MAX_STATION_NUM] OF INT := [0];
	iWaitedCycleCount: INT := 0;
	xForceAxisOff: BOOL;(*强制下伺服标志*)
	xFlag_AllInchRun_ing: BOOL;
	iMotionModePrn : INT;//版辊运动模式
						//0、电子齿轮
						//1、点位 --恢复相位等
						//2、Jog模式
	astStTStGearParam: ARRAY [1..MAX_STATION_NUM] OF TStGearParam;
	fbKS_FB_SyncAxisParam_Trap : KS_FB_SyncAxisParam_Trap;
	xKeepServo: BOOL;//保持伺服标志

	afbTRIG_Start_Servo: ARRAY [1..MAX_STATION_NUM] OF R_TRIG;
	afbTRIG_Stop_Servo: ARRAY [1..MAX_STATION_NUM] OF R_TRIG;
	axServoOn: ARRAY [1..MAX_STATION_NUM] OF BOOL;

	iN: INT;

	iRtn_McMulFun : INT ;
	iRtn_McMulFun_Pre : INT ;
	sTMultiMcFunctionReadPrm : TMultiMcFunctionReadPrm;
	alrVarValue : ARRAY [1..80] OF LREAL;

	//2026.01.28.173520 | + | 横向伺服控制
	fbKS_FB_AxisPosCtl_Trap : KS_FB_AxisPosCtl_Trap;
	alrTarp_EncPos						: ARRAY [1..MAX_UNIT_NUM] OF LREAL;//横向点位轴的编码器位置

	aiWaitingModalChange : ARRAY [1..MAX_STATION_NUM] OF INT;

	//2026.04.02.91845 新增

	iUnitId: INT;
	iTypeId: INT;
	iCoreId: INT;
	iAxisId: INT;
	iGroupId : INT;
	iAdjAxisId : INT;
END_VAR

{IMPLEMENTATION}
IF i_xEn THEN
	IF i_pstStSysParam<>0 AND i_pastStSetPrm <> 0 AND i_pastStGetMotionSts <> 0 AND
		i_pastStMotorParam_Trap <> 0 AND i_pstStHYLogFifo <> 0 AND i_pastStIOMap_Main_FE <> 0 AND i_pastStIOMap_Axis_FE <> 0 THEN
(*这里作为同步使能、速度等参数*)

		fbKS_FB_SyncAxisParam_Trap(
			i_xEn:= TRUE,
			i_iGrpId:= i_iGrpId,
			i_iGrpUnitNum_Pu:= i_iGrpUnitNum_Pu,
			i_aiGrpUnitList:= i_aiGrpUnitList,
			i_iGrpTrapMotion_Num:= i_iGrpTrapMotion_Num,
			i_aiGrpTrapMotion_StdList:= i_aiGrpTrapMotion_StdList,
			i_pstStSysParam:= i_pstStSysParam,
			i_pastStMotorParam_Trap := i_pastStMotorParam_Trap,
			i_pstStSysStationInf := i_pstStSysStationInf,
			i_pstStSysGantryAxisInf := i_pstStSysGantryAxisInf,
			i_pastStGetMotionSts := i_pastStGetMotionSts,
			i_palrTarp_EncPos := ADR(alrTarp_EncPos)
		);

		fbKS_FB_AxisPosCtl_Trap(
			i_xEn:= TRUE,
			i_iGrpId:= i_iGrpId,
			i_iGrpUnitNum_Pu:= i_iGrpUnitNum_Pu,
			i_aiGrpUnitList:= i_aiGrpUnitList,
			i_iGrpTrapMotion_Num:= i_iGrpTrapMotion_Num,
			i_aiGrpTrapMotion_StdList:= i_aiGrpTrapMotion_StdList,
			i_pstStSysParam:= i_pstStSysParam,
			i_pastStMotorParam_Trap:= i_pastStMotorParam_Trap,
			i_xHorManuCtrl:= i_xHorManuCtrl,
			i_alrTarp_EncPos:= alrTarp_EncPos,
			i_pastStIOMap_AxisBasic:= i_pastStIOMap_Axis_FE,
			i_pastStAxisRapidAdjProf_H:= i_pastStAxisRapidAdjProf_H,
			i_paxLimit_Left_Wr:= i_paxLimit_Left_Wr,
			i_paxLimit_Right_Wr:= i_paxLimit_Right_Wr,
			i_paxLimit_Left_WrClr:= i_paxLimit_Left_WrClr,
			i_paxLimit_Right_WrClr:= i_paxLimit_Right_WrClr,
			i_pastStGetMotionSts:=i_pastStGetMotionSts,
			i_pstStSysStationInf:=i_pstStSysStationInf,
			i_pstStSysGantryAxisInf :=i_pstStSysGantryAxisInf,
			i_pastStAxisIdListInf :=i_pastStAxisIdListInf,
);

		pstStGrpParam_Save := ADR(i_pstStSysParam^.astStGrpParam_Save[i_iGrpId]);
		pstStGrpParam_UnSave := ADR(i_pstStSysParam^.astStGrpParam_UnSave[i_iGrpId]);

		FOR iN:=1 TO i_iGrpTrapMotion_Num BY 1 DO
			afbTRIG_Start_Servo[iN](CLK:= i_pastStMotorParam_Trap^[iN].xMoveEn);
			afbTRIG_Stop_Servo[iN](CLK:= NOT i_pastStMotorParam_Trap^[iN].xMoveEn);

			IF afbTRIG_Start_Servo[iN].Q THEN
				IF i_pastStMotorParam_Trap^[iN].iMoveStep= MOTION_STEP_Nothing THEN
					i_pastStMotorParam_Trap^[iN].iMoveStep:= MOTIONCTL_STEP_SETMOTIONMODE;
				ELSE;
				END_IF
			END_IF
			IF afbTRIG_Stop_Servo[iN].Q THEN
				IF i_pastStMotorParam_Trap^[iN].iMoveStep= MOTION_STEP_Nothing OR
					i_pastStMotorParam_Trap^[iN].iMoveStep= MOTIONCTL_STEP_AXISOFF THEN
					;
				ELSE
					i_pastStMotorParam_Trap^[iN].iMoveStep:= MOTIONCTL_STEP_AXISOFF;
				END_IF
			END_IF

			CASE i_pastStMotorParam_Trap^[iN].iMoveStep OF
			MOTION_STEP_Nothing:
				;
			MOTIONCTL_STEP_AXISOFF:
				iRtn:= KS_SetMotionServoOff(
					i_iAxisId:= i_pastStMotorParam_Trap^[iN].iAxisId,
					i_iCoreId:= i_pastStMotorParam_Trap^[iN].iCoreId,
					i_iStationId:= i_pastStMotorParam_Trap^[iN].iStationId,
					i_xForceAxisOff:= FALSE,
					i_dwMotionSts:= i_pastStGetMotionSts^[i_pastStMotorParam_Trap^[iN].iAxisId].dwMotionSts,
					i_dwDriverSts:= i_pastStGetMotionSts^[i_pastStMotorParam_Trap^[iN].iAxisId].dwDriverSts,
					i_pxServoOn:= ADR(axServoOn[iN]),
					i_pstStHYLogFifo:= i_pstStHYLogFifo);

				IF iRtn<>0 THEN
					IF aiRetryCount[iN]>=iMaxRetryTimes THEN(*如果失败次数超过3次则就结束绝对位置确认这个操作*)
						i_pastStMotorParam_Trap^[iN].iMoveStep:= MOTIONCTL_STEP_AXISOFF;
					ELSE
						aiRetryCount[iN]:= aiRetryCount[iN]+1;
					END_IF
				ELSE
					aiRetryCount[iN]:= 0;
					i_pastStMotorParam_Trap^[iN].iMoveStep:= MOTION_STEP_Nothing;
				END_IF

				//2025.10.27.164954 | bai.zy |
				i_pastStSetPrm^[i_pastStMotorParam_Trap^[iN].iAxisId].prm.trapPrm.axis_ctrl:= 2;
			MOTIONCTL_STEP_SETMOTIONMODE:
				iRtn:= KS_SetMotionMode(
					i_iAxisId:= i_pastStMotorParam_Trap^[iN].iAxisId,
					i_iCoreId:= i_pastStMotorParam_Trap^[iN].iCoreId,
					i_iStationId:= i_pastStMotorParam_Trap^[iN].iStationId,
					i_iMoveMode:= 2,
					i_iAxisId_Master:= 64,
					i_xMasterType := FALSE,
					i_pstStHYLogFifo:= i_pstStHYLogFifo);
				IF iRtn<>0 THEN
					IF aiRetryCount[iN]>=iMaxRetryTimes THEN(*如果失败次数超过3次则就结束绝对位置确认这个操作*)
						i_pastStMotorParam_Trap^[iN].iMoveStep:= MOTIONCTL_STEP_AXISOFF;
					ELSE
						aiRetryCount[iN]:= aiRetryCount[iN]+1;
					END_IF
				ELSE
					aiRetryCount[iN]:= 0;
					i_pastStMotorParam_Trap^[iN].iMoveStep:= MOTIONCTL_STEP_CLRSTS;
				END_IF
			MOTIONCTL_STEP_CLRSTS:
				iRtn:= KS_SetMotionClrSts(
					i_iAxisId:= i_pastStMotorParam_Trap^[iN].iAxisId,
					i_iCoreId:= i_pastStMotorParam_Trap^[iN].iCoreId,
					i_iStationId:= i_pastStMotorParam_Trap^[iN].iStationId,
					i_pstStHYLogFifo:= i_pstStHYLogFifo);
				IF iRtn<>0 THEN
					IF aiRetryCount[iN]>=iMaxRetryTimes THEN(*如果失败次数超过3次则就结束绝对位置确认这个操作*)
						i_pastStMotorParam_Trap^[iN].iMoveStep:= MOTIONCTL_STEP_AXISOFF;
					ELSE
						aiRetryCount[iN]:= aiRetryCount[iN]+1;
					END_IF
				ELSE
					aiRetryCount[iN]:= 0;
					i_pastStMotorParam_Trap^[iN].iMoveStep:= MOTIONCTL_STEP_AXISON;
				END_IF
			MOTIONCTL_STEP_AXISON:
				iRtn:= KS_SetMotionServoOn(
					i_iAxisId:= i_pastStMotorParam_Trap^[iN].iAxisId,
					i_iCoreId:= i_pastStMotorParam_Trap^[iN].iCoreId,
					i_iStationId:= i_pastStMotorParam_Trap^[iN].iStationId,
					i_pxMoveEn := ADR(i_pastStMotorParam_Trap^[iN].xMoveEn),
					i_pxServoOn:= ADR(axServoOn[iN]),
					i_pstStHYLogFifo:= i_pstStHYLogFifo);
				IF iRtn<>0 THEN
					IF aiRetryCount[iN]>=iMaxRetryTimes THEN(*如果失败次数超过3次则就结束绝对位置确认这个操作*)
						i_pastStMotorParam_Trap^[iN].iMoveStep:= MOTIONCTL_STEP_AXISOFF;
					ELSE
						aiRetryCount[iN]:= aiRetryCount[iN]+1;
					END_IF
				ELSE
					aiRetryCount[iN]:= 0;
					i_pastStMotorParam_Trap^[iN].iMoveStep:= MOTIONCTL_STEP_WaitingModalChanged;
				END_IF

			MOTIONCTL_STEP_WaitingModalChanged:
				aiWaitingModalChange[iN] := aiWaitingModalChange[iN] + 1;
				IF aiWaitingModalChange[iN] > 50 THEN
					aiWaitingModalChange[iN] := 0;
					i_pastStMotorParam_Trap^[iN].iMoveStep:= MOTIONCTL_STEP_CHECKAXISON;
				END_IF
			MOTIONCTL_STEP_CHECKAXISON:
				iRtn:= KS_SetMotionCheckServoOn(
					i_iAxisId:= i_pastStMotorParam_Trap^[iN].iAxisId,
					i_iCoreId:= i_pastStMotorParam_Trap^[iN].iCoreId,
					i_iStationId:= i_pastStMotorParam_Trap^[iN].iStationId,
					i_pxMoveEn := ADR(i_pastStMotorParam_Trap^[iN].xMoveEn),
					i_dwMotionSts:= i_pastStGetMotionSts^[i_pastStMotorParam_Trap^[iN].iAxisId].dwMotionSts,
					i_dwDriverSts:= i_pastStGetMotionSts^[i_pastStMotorParam_Trap^[iN].iAxisId].dwDriverSts,
					i_pxServoOn:= ADR(axServoOn[iN]),
					i_pstStHYLogFifo:= i_pstStHYLogFifo);
				IF iRtn<>0 THEN
					IF aiRetryCount[iN]>=iMaxRetryTimes THEN(*如果失败次数超过3次则就结束绝对位置确认这个操作*)
						i_pastStMotorParam_Trap^[iN].iMoveStep:= MOTIONCTL_STEP_AXISOFF;
						axServoOn[iN] := FALSE;
					ELSE
						aiRetryCount[iN]:= aiRetryCount[iN]+1;
					END_IF
				ELSE
					aiRetryCount[iN]:= 0;
					i_pastStMotorParam_Trap^[iN].iMoveStep:= MOTIONCTL_STEP_WRITEDATA_Run;
				END_IF
			MOTIONCTL_STEP_WRITEDATA_Run:
				i_pastStSetPrm^[iN].profileMode := 1;
				i_pastStSetPrm^[iN].prm.trapPrm.axis_ctrl:= 3;
				i_pastStSetPrm^[iN].prm.trapPrm.axis_id:= INT_TO_UINT(i_pastStMotorParam_Trap^[iN].iAxisId);
				i_pastStSetPrm^[iN].prm.trapPrm.axis_mode:= 1;
				i_pastStSetPrm^[iN].prm.trapPrm.reserve:= 0;
				i_pastStSetPrm^[iN].prm.trapPrm.reserve2[1]:= 0;
				i_pastStSetPrm^[iN].prm.trapPrm.reserve2[2]:= 0;
				i_pastStSetPrm^[iN].prm.trapPrm.target_pos:= i_pastStMotorParam_Trap^[iN].liTargetPos;
				i_pastStSetPrm^[iN].prm.trapPrm.max_vel:= i_pastStMotorParam_Trap^[iN].udiTargetVel;
			END_CASE
		END_FOR

		(*2.大指令写*)
		sTMultiMcFunctionReadPrm.readCommandVarTableIndex := 1;
		sTMultiMcFunctionReadPrm.readCount := 0;
		sTMultiMcFunctionReadPrm.pVarValue := ADR(alrVarValue);
		dwRtn:= SysMemCmp(i_pastStSetPrm,ADR(astStSetPrm_Pre),SIZEOF(astStSetPrm_Pre));
		IF dwRtn<>0 THEN
			iRtn_McMulFun:=GTN_StartMcMultiFunction(1,INT_TO_UINT(i_iGrpTrapMotion_Num),1,i_pastStSetPrm,ADR(sTMultiMcFunctionReadPrm));
			IF iRtn_McMulFun <> 0 AND iRtn_McMulFun_Pre <> iRtn_McMulFun THEN
				KS_HY_AddMsgToLog(g_pstStHYLogFifo, LOG_LEVEL_ALARM, 'GTN_StartMcMultiFunction Trap Err!', INT_TO_STRING(iRtn_McMulFun));
			END_IF
			iRtn_McMulFun_Pre := iRtn_McMulFun;
		END_IF
		SysMemCpy(ADR(astStSetPrm_Pre),i_pastStSetPrm,SIZEOF(i_pastStSetPrm^));

		//2026.04.02.92001 新增拿横向编码器 Hou.N
			FOR iN := 1 TO  i_iGrpTrapMotion_Num BY 1 DO
				KS_GetAxisIdForMotByStation_V2(
					i_iStationId:= i_aiGrpTrapMotion_StdList[iN],
					i_piAxisId:= ADR(iAxisId),
					i_piTypeId:= ADR(iTypeId),
					i_piUnitId:= ADR(iUnitId),
					i_piCoreId:= ADR(iCoreId),
					i_piGroupId:= ADR(iGroupId),
					i_piAdjAxisId:= ADR(iAdjAxisId),
					i_pstStSysStationInf:= i_pstStSysStationInf);
				IF iTypeId= TYPE_UNIT_HORIZ THEN
					g_alrTrap_EncPos[iUnitId]	:= i_pastStGetMotionSts^[iAxisId].lrPos_Enc;
					g_arTrapPos_mm[iUnitId]:=	g_alrTrap_EncPos[iUnitId]*
												i_pstStSysParam^.astStUnitParam_Save[iUnitId].rScrewPitch_Horz*
												UINT_TO_REAL(i_pstStSysParam^.astStUnitParam_Save[iUnitId].uiDen_Horz)
												/GC_LRMOTORPPR_TRAP/UINT_TO_REAL(i_pstStSysParam^.astStUnitParam_Save[iUnitId].uiNum_Horz);
				END_IF
			END_FOR

	ELSE;
	END_IF
ELSE
	;
END_IF

(* ---- KS_FB_SyncAxisParam_Trap.st ---- *)
(*@CES
Name=KS_FB_SyncAxisParam_Trap
Type=FunctionBlock
TypeGuid=6f9dac99-8de1-4efc-8465-68ac443b7d08
Guid=6588b639-e838-4495-9484-0472b9b3fcb8
HasDeclaration=True
HasImplementation=True
*)
{DECLARATION}
FUNCTION_BLOCK KS_FB_SyncAxisParam_Trap
VAR_INPUT
	i_xEn: BOOL;
	i_iGrpId: INT;
	i_iGrpUnitNum_Pu : INT;
	i_aiGrpUnitList: ARRAY [1..MAX_UNIT_NUM] OF INT;
	i_iGrpTrapMotion_Num: INT;
	i_aiGrpTrapMotion_StdList: ARRAY [1..MAX_STATION_NUM] OF INT;

	i_pstStSysParam: POINTER TO StSysParam;
	i_pastStMotorParam_Trap: POINTER TO ARRAY [1..MAX_STATION_NUM] OF StMotorParam_Trap;

	i_pstStSysStationInf			:POINTER TO StSysStationInf;
	i_pstStSysGantryAxisInf : POINTER TO StSysGantryAxisInf;
	i_pastStGetMotionSts: POINTER TO ARRAY [1..MAX_STATION_NUM] OF StGetMotionSts;
	i_palrTarp_EncPos		:POINTER TO ARRAY [1..MAX_UNIT_NUM] OF LREAL;//横向点位轴的编码器位置

END_VAR
VAR_OUTPUT
END_VAR
VAR
	iRtn : INT;
	iN: INT;
	iUnitId: INT;
	iTypeId: INT;
	iCoreId: INT;
	iAxisId: INT;
	iGroupId : INT;
	iAdjAxisId : INT;
	pstStGrpParam_Save: POINTER TO StGrpParam_Save;
	pstStGrpParam_UnSave: POINTER TO StGrpParam_UnSave;

	xInit_TrapPoint : BOOL;
	iAxisCount : INT;
	aiTargetStation : ARRAY [1..MAX_STATION_NUM] OF INT;//压力电机站列表
	aliABSEncPos : ARRAY [1..MAX_STATION_NUM] OF LINT;//零位绝对编码器位置
	axAxisRev : ARRAY [1..MAX_STATION_NUM] OF BOOL;//零位绝对编码器位置
END_VAR

{IMPLEMENTATION}
IF i_xEn THEN
	IF i_pstStSysParam<>0 AND i_pastStMotorParam_Trap <> 0 AND
		i_pstStSysStationInf <> 0 AND i_pstStSysGantryAxisInf <> 0 THEN

		FOR iN:=1 TO i_iGrpUnitNum_Pu BY 1 DO
			iUnitId:= i_aiGrpUnitList[iN];
		(*横向电机方向*)
			i_pstStSysParam^.astStUnitParam_UnSave[iUnitId].xMotRev_Horiz_:=
					i_pstStSysParam^.stStSysParam_UnSave.stStSysCfgStruct.astStAxisCfgStruct_HORIZ_[iUnitId].dwAxisProf.1;
		(*横向减速比*)
			i_pstStSysParam^.astStUnitParam_Save[iUnitId].uiNum_Horz:=
					i_pstStSysParam^.astStGrpParam_Save[i_iGrpId].uiNum_Horz;
			i_pstStSysParam^.astStUnitParam_Save[iUnitId].uiDen_Horz:=
					i_pstStSysParam^.astStGrpParam_Save[i_iGrpId].uiDen_Horz;
			i_pstStSysParam^.astStUnitParam_Save[iUnitId].rScrewPitch_Horz:=
					i_pstStSysParam^.astStGrpParam_Save[i_iGrpId].rScrewPitch_Horz;
		END_FOR

		FOR iN:=1 TO i_iGrpTrapMotion_Num BY 1 DO
			KS_GetAxisIdForMotByStation_V2(
					i_iStationId:= i_aiGrpTrapMotion_StdList[iN],
					i_piAxisId:= ADR(iAxisId),
					i_piTypeId:= ADR(iTypeId),
					i_piUnitId:= ADR(iUnitId),
					i_piCoreId:= ADR(iCoreId),
					i_piGroupId:= ADR(iGroupId),
					i_piAdjAxisId:= ADR(iAdjAxisId),
					i_pstStSysStationInf:= i_pstStSysStationInf);

			CASE iTypeId OF
			TYPE_UNIT_HORIZ:
				i_pastStMotorParam_Trap^[iUnitId].iAxisId := iAxisId;
				i_pastStMotorParam_Trap^[iUnitId].iCoreId := iCoreId;
				i_pastStMotorParam_Trap^[iUnitId].iStationId := i_aiGrpTrapMotion_StdList[iN];
				i_pastStMotorParam_Trap^[iUnitId].iUnitId := iUnitId;
				i_pastStMotorParam_Trap^[iUnitId].xMoveRev := i_pstStSysParam^.astStUnitParam_UnSave[iUnitId].xMotRev_Horiz_;
				i_pastStMotorParam_Trap^[iUnitId].uiAxisNum := i_pstStSysParam^.astStUnitParam_Save[iUnitId].uiNum_PrnRoller_Pressure;
				i_pastStMotorParam_Trap^[iUnitId].uiAxisDen := i_pstStSysParam^.astStUnitParam_Save[iUnitId].uiDen_PrnRoller_Pressure;
				i_pastStMotorParam_Trap^[iUnitId].rScrewPitch_ := i_pstStSysParam^.astStUnitParam_Save[iUnitId].rScrewPitch_PrnRoller_Pressure;
				i_pastStMotorParam_Trap^[iUnitId].xMoveEn := g_xMoveEnTrap;//2026.01.28.115155 | + | 点位运动一直维持使能，后续还是要增加标志

				i_palrTarp_EncPos^[iUnitId] := i_pastStGetMotionSts^[iAxisId].lrPos_Enc;
			END_CASE
		END_FOR

		IF NOT xInit_TrapPoint THEN
			FOR iN := 1 TO  i_iGrpTrapMotion_Num BY 1 DO
				KS_GetAxisIdForMotByStation_V2(
					i_iStationId:= i_aiGrpTrapMotion_StdList[iN],
					i_piAxisId:= ADR(iAxisId),
					i_piTypeId:= ADR(iTypeId),
					i_piUnitId:= ADR(iUnitId),
					i_piCoreId:= ADR(iCoreId),
					i_piGroupId:= ADR(iGroupId),
					i_piAdjAxisId:= ADR(iAdjAxisId),
					i_pstStSysStationInf:= i_pstStSysStationInf);

				IF iTypeId= TYPE_UNIT_HORIZ THEN
					iAxisCount := iAxisCount + 1;
					aiTargetStation[iAxisCount] := (i_aiGrpTrapMotion_StdList[iN]);
					aliABSEncPos[iAxisCount]:= i_pstStSysParam^.astStRSV_UnitParam_Save[iUnitId].liABSPos_Trap;//g_aliABSPos_Horiz[iUnitId];
					axAxisRev[iAxisCount]:=i_pstStSysParam^.astStUnitParam_UnSave[iUnitId].xMotRev_Horiz_;

					iRtn := KS_SetTrapDir(
						i_xEn:= TRUE,
						i_iAxisId:= iAxisId,
						i_iCoreId:= iCoreId,
						i_xRevDir:= axAxisRev[iAxisCount]);
				END_IF
			END_FOR

			iRtn := KS_SetTrapCoordinate(
						i_xEn:= TRUE,
						i_iTarget_Num:= iAxisCount,
						i_paiTargetStationList:= ADR(aiTargetStation),
						i_paliABSEncPos:= ADR(aliABSEncPos),
						i_paxAxisRev:= ADR(axAxisRev),
						i_pastStAxisIdListInf:= ADR(g_astStAxisIdListInf),
						i_pastStGetMotionSts:= ADR(g_astStGetMotionSts),
						i_pstStSysStationInf := i_pstStSysStationInf,
						i_pstStSysGantryAxisInf := i_pstStSysGantryAxisInf,
						ADR(g_alrCurrentAbsPos_Trap));
			xInit_TrapPoint := TRUE;
		END_IF
	ELSE;
	END_IF
ELSE
	;
END_IF
